     ELSIF (#statErrorAutoCleared = FALSE AND NOT #tempExecute) AND (#statErrorUserCleared = FALSE) AND (#statError = TRUE) THEN
       REGION after user/auto cleared 
         // if autocleared error is acknowledged
         #statValid := TRUE;
         #statBusy := FALSE;
         #statError := FALSE;
         #statDiagnostics.status := #STATUS_READY;
       END_REGION after user/auto cleared or command aborted
     END_IF;

     REGION Write static values to outputs
       #valid := #statValid;
       #done := #statDone;
       #busy := #statBusy;
       #error := #statError;
       #status := #statDiagnostics.status;
       // if ENO mechanism is not used / not wanted replace the following line by --> ENO := TRUE;
       ENO := NOT #statError;
     END_REGION Write static values to outputs
   END_REGION
END_FUNCTION_BLOCK